      FC_W[1,12] := 0.07566059;
      FC_W[1,13] := 0.35968998;
      FC_W[1,14] := -0.17466193;
      FC_W[1,15] := 1.00617445;
      FC_W[1,16] := 0.29971626;
      FC_W[1,17] := -0.15427162;
      FC_W[1,18] := 0.06198071;
      FC_W[1,19] := 0.48209724;
      FC_W[1,20] := -1.77777910;
      FC_W[1,21] := 0.30678549;
      FC_W[1,22] := -0.06820694;
      FC_W[1,23] := -1.06389523;
      FC_W[1,24] := 1.40704405;
      FC_W[1,25] := 0.86564183;
      FC_W[1,26] := 0.86175865;
      FC_W[1,27] := -0.30832738;
      FC_W[1,28] := 0.12632002;
      FC_W[1,29] := 0.22659495;
      FC_W[1,30] := -0.13902418;
      FC_W[1,31] := -0.99291939;
      FC_W[2,0] := 0.04160358;
      FC_W[2,1] := 0.28197494;
      FC_W[2,2] := -0.02089060;
      FC_W[2,3] := 0.47015443;
      FC_W[2,4] := 0.34037617;
      FC_W[2,5] := -0.41242811;
      FC_W[2,6] := -0.82493418;
      FC_W[2,7] := 0.78098351;
      FC_W[2,8] := -0.39970401;
      FC_W[2,9] := 1.02419770;
      FC_W[2,10] := -0.33057141;
      FC_W[2,11] := 0.13100362;
      FC_W[2,12] := -1.50004947;
      FC_W[2,13] := -0.18024392;
      FC_W[2,14] := 0.19656396;
      FC_W[2,15] := -1.08431160;
      FC_W[2,16] := -0.22757976;
      FC_W[2,17] := -0.09310954;
      FC_W[2,18] := 1.20083344;
      FC_W[2,19] := -0.90194166;
      FC_W[2,20] := 0.46690372;
      FC_W[2,21] := -0.28373122;
      FC_W[2,22] := 0.44820097;
      FC_W[2,23] := 1.57939780;
      FC_W[2,24] := -0.41811836;
      FC_W[2,25] := 0.45971355;
      FC_W[2,26] := -0.05362111;
      FC_W[2,27] := -0.62090284;
      FC_W[2,28] := -0.41635084;
      FC_W[2,29] := 1.19535244;
      FC_W[2,30] := 0.22620986;
      FC_W[2,31] := -0.29096127;
      FC_W[3,0] := 0.69258898;
      FC_W[3,1] := -0.10189002;
      FC_W[3,2] := -0.35127911;
      FC_W[3,3] := -0.06208733;
      FC_W[3,4] := -0.31526309;
      FC_W[3,5] := -0.58414000;
      FC_W[3,6] := 0.04904716;
      FC_W[3,7] := 0.37988806;
      FC_W[3,8] := -0.33488220;
      FC_W[3,9] := 0.67849815;
      FC_W[3,10] := 0.02032584;
      FC_W[3,11] := -0.11450892;
      FC_W[3,12] := 0.75389469;
      FC_W[3,13] := -0.00020683;
      FC_W[3,14] := 0.11827329;
      FC_W[3,15] := 0.03889267;
      FC_W[3,16] := 0.17466927;
      FC_W[3,17] := -0.05837984;
      FC_W[3,18] := 0.16143340;
      FC_W[3,19] := -0.25548884;
      FC_W[3,20] := 0.36278751;
      FC_W[3,21] := 0.31648728;
      FC_W[3,22] := -0.78370738;
      FC_W[3,23] := -0.28512084;
      FC_W[3,24] := -0.33843708;
      FC_W[3,25] := 0.04330043;
      FC_W[3,26] := -0.25837252;
      FC_W[3,27] := 0.40221891;
      FC_W[3,28] := 0.07115368;
      FC_W[3,29] := 1.57388341;
      FC_W[3,30] := 0.08364432;
      FC_W[3,31] := 0.69666040;
      FC_W[4,0] := 0.17098659;
      FC_W[4,1] := 0.70854473;
      FC_W[4,2] := 0.32589009;
      FC_W[4,3] := -0.19657923;
      FC_W[4,4] := 0.02836942;
      FC_W[4,5] := -0.33067968;
      FC_W[4,6] := -0.28083199;
      FC_W[4,7] := 0.21882291;
      FC_W[4,8] := 0.44031367;
      FC_W[4,9] := -0.08098698;
      FC_W[4,10] := 0.40485817;
      FC_W[4,11] := -0.28698298;
      FC_W[4,12] := 0.25233796;
      FC_W[4,13] := -0.10523839;
      FC_W[4,14] := -0.44006598;
      FC_W[4,15] := -0.39039072;
      FC_W[4,16] := 0.15023036;
      FC_W[4,17] := 0.09987778;
      FC_W[4,18] := -0.55138695;
      FC_W[4,19] := 0.97002214;
      FC_W[4,20] := -1.32036424;
      FC_W[4,21] := 0.12111247;
      FC_W[4,22] := 0.17146327;
      FC_W[4,23] := -0.14426313;
      FC_W[4,24] := -1.44331551;
      FC_W[4,25] := -0.32387802;
      FC_W[4,26] := -0.86985487;
      FC_W[4,27] := 0.16190216;
      FC_W[4,28] := -0.25917780;
      FC_W[4,29] := 0.87935007;
      FC_W[4,30] := -0.04532806;
      FC_W[4,31] := 0.12371654;
      FC_W[5,0] := 0.16069181;
      FC_W[5,1] := 1.64132881;
      FC_W[5,2] := 0.09314496;
      FC_W[5,3] := 0.30746382;
      FC_W[5,4] := -0.44713461;
      FC_W[5,5] := -0.17269248;
      FC_W[5,6] := -0.43764487;
      FC_W[5,7] := -0.55917907;
      FC_W[5,8] := 0.07907125;
      FC_W[5,9] := 0.32444280;
      FC_W[5,10] := 0.17686915;
      FC_W[5,11] := -0.43060029;
      FC_W[5,12] := -0.11524609;
      FC_W[5,13] := -0.43634474;
      FC_W[5,14] := -0.84067672;
      FC_W[5,15] := 0.12469457;
      FC_W[5,16] := 0.36836424;
      FC_W[5,17] := -0.39146784;
      FC_W[5,18] := 0.77493954;
      FC_W[5,19] := -0.39445737;
      FC_W[5,20] := 0.13570420;
      FC_W[5,21] := -0.30796599;
      FC_W[5,22] := 0.57390678;
      FC_W[5,23] := -0.10128630;
      FC_W[5,24] := 0.46898919;
      FC_W[5,25] := -0.44309253;
      FC_W[5,26] := 0.08969644;
      FC_W[5,27] := -0.19782862;
      FC_W[5,28] := 2.73940182;
      FC_W[5,29] := 0.16153421;
      FC_W[5,30] := -0.12013239;
      FC_W[5,31] := -0.56593496;
      FC_W[6,0] := -0.57114196;
      FC_W[6,1] := 1.38476813;
      FC_W[6,2] := 1.11997521;
      FC_W[6,3] := 0.02632367;
      FC_W[6,4] := -0.45034066;
      FC_W[6,5] := 1.03288424;
      FC_W[6,6] := -0.40567783;
      FC_W[6,7] := 0.16608752;
      FC_W[6,8] := 0.03270433;
      FC_W[6,9] := -0.35795641;
      FC_W[6,10] := 0.00975101;
      FC_W[6,11] := -0.41937128;
      FC_W[6,12] := -0.19609804;
      FC_W[6,13] := -0.28889647;
      FC_W[6,14] := -0.96404856;
      FC_W[6,15] := 0.08155423;
      FC_W[6,16] := 0.09745946;
      FC_W[6,17] := 0.17013049;
      FC_W[6,18] := 0.17057557;
      FC_W[6,19] := -0.79009062;
      FC_W[6,20] := 0.26148456;
      FC_W[6,21] := -0.41126329;
      FC_W[6,22] := -0.92280918;
      FC_W[6,23] := -0.19497190;
      FC_W[6,24] := 0.56321335;
      FC_W[6,25] := -0.69397563;
      FC_W[6,26] := -0.11093070;
      FC_W[6,27] := -0.12486640;
      FC_W[6,28] := -0.51809597;
      FC_W[6,29] := 0.44581598;
      FC_W[6,30] := -0.07224379;
      FC_W[6,31] := 0.58158380;
      FC_W[7,0] := 0.41476303;
      FC_W[7,1] := -0.03894622;
      FC_W[7,2] := -0.50756085;
      FC_W[7,3] := -0.26348099;
      FC_W[7,4] := 0.08712668;
      FC_W[7,5] := -0.37651458;
      FC_W[7,6] := 0.26482788;
      FC_W[7,7] := -0.29581240;
      FC_W[7,8] := 0.05395310;
      FC_W[7,9] := 0.41241437;
      FC_W[7,10] := -0.15156971;
      FC_W[7,11] := 0.26749688;
      FC_W[7,12] := 0.97054368;
      FC_W[7,13] := -0.03540496;
      FC_W[7,14] := -0.09778718;
      FC_W[7,15] := -0.39193475;
      FC_W[7,16] := -0.01532598;
      FC_W[7,17] := -0.11887385;
      FC_W[7,18] := -0.30799413;
      FC_W[7,19] := -0.20951317;
      FC_W[7,20] := 0.46884289;
      FC_W[7,21] := 0.08239307;
      FC_W[7,22] := -0.41243985;
      FC_W[7,23] := -0.14386208;
      FC_W[7,24] := -0.56366146;
      FC_W[7,25] := 0.05347069;
      FC_W[7,26] := -0.06422243;
      FC_W[7,27] := -0.14232105;
      FC_W[7,28] := 0.08967300;
      FC_W[7,29] := 2.09215212;
      FC_W[7,30] := -0.41609016;
      FC_W[7,31] := 0.61930108;
      FC_W[8,0] := 0.41138357;
      FC_W[8,1] := -0.13876545;
      FC_W[8,2] := -0.47696707;
      FC_W[8,3] := -0.58067173;
      FC_W[8,4] := -0.76539934;
      FC_W[8,5] := -0.48228866;
      FC_W[8,6] := 0.25288635;
      FC_W[8,7] := 1.26393640;
      FC_W[8,8] := -0.18708183;
      FC_W[8,9] := 1.05916786;
      FC_W[8,10] := -0.21405555;
      FC_W[8,11] := -0.73763049;
      FC_W[8,12] := -0.49388906;
      FC_W[8,13] := 0.23774624;
      FC_W[8,14] := 0.03641314;
      FC_W[8,15] := 0.43136188;
      FC_W[8,16] := -0.34853166;
      FC_W[8,17] := 0.45351282;
      FC_W[8,18] := 0.12007232;
      FC_W[8,19] := -0.09311971;
      FC_W[8,20] := 0.10139518;
      FC_W[8,21] := 0.13798890;
      FC_W[8,22] := -0.75192511;
      FC_W[8,23] := -0.33668301;
      FC_W[8,24] := 0.14659424;
      FC_W[8,25] := -0.00453089;
      FC_W[8,26] := -0.35082975;
      FC_W[8,27] := 0.47500724;
      FC_W[8,28] := 0.02143906;
      FC_W[8,29] := 0.81066149;
      FC_W[8,30] := 0.42516547;
      FC_W[8,31] := 1.48935926;
      FC_W[9,0] := 0.29422590;
      FC_W[9,1] := -0.02413537;
      FC_W[9,2] := -0.57707560;
      FC_W[9,3] := -0.44330636;
      FC_W[9,4] := -0.02986326;
      FC_W[9,5] := -0.32138100;
      FC_W[9,6] := 0.33747303;
      FC_W[9,7] := -0.02603977;
      FC_W[9,8] := 0.16214876;
      FC_W[9,9] := 0.54148763;
      FC_W[9,10] := -0.23998420;
      FC_W[9,11] := 0.06466576;
      FC_W[9,12] := 0.47260144;
      FC_W[9,13] := 0.04922871;
      FC_W[9,14] := -0.13990949;
      FC_W[9,15] := -0.24958028;
      FC_W[9,16] := -0.20513535;
      FC_W[9,17] := 0.11604570;
      FC_W[9,18] := -0.38338530;
      FC_W[9,19] := -0.16188677;
      FC_W[9,20] := 0.37325716;
      FC_W[9,21] := -0.01747377;
      FC_W[9,22] := -0.37153879;
      FC_W[9,23] := -0.15362059;
      FC_W[9,24] := -0.37243831;
      FC_W[9,25] := 0.01588886;
      FC_W[9,26] := -0.08001896;
      FC_W[9,27] := -0.14023392;
      FC_W[9,28] := 0.07176708;
      FC_W[9,29] := 1.81881726;
      FC_W[9,30] := -0.30937484;
      FC_W[9,31] := 0.93038040;
      FC_W[10,0] := -0.05140001;
      FC_W[10,1] := -0.21192010;
      FC_W[10,2] := -0.34014732;
      FC_W[10,3] := -0.41698745;
      FC_W[10,4] := 1.15412712;
      FC_W[10,5] := -0.76638728;
      FC_W[10,6] := -0.36194009;
      FC_W[10,7] := -0.14446546;
      FC_W[10,8] := 0.05265777;
      FC_W[10,9] := 0.60072738;
      FC_W[10,10] := 0.43118945;
      FC_W[10,11] := 0.83294547;
      FC_W[10,12] := 0.67825025;
      FC_W[10,13] := 0.19051756;
      FC_W[10,14] := 1.69663048;
      FC_W[10,15] := -0.22305325;
      FC_W[10,16] := -0.32500228;
      FC_W[10,17] := 0.31870443;
      FC_W[10,18] := 0.10095058;
      FC_W[10,19] := -0.75147802;
      FC_W[10,20] := -0.45519939;
      FC_W[10,21] := 0.01013143;
      FC_W[10,22] := 0.00206094;
      FC_W[10,23] := 0.25191501;
      FC_W[10,24] := 0.39815706;
      FC_W[10,25] := -0.34215525;
      FC_W[10,26] := -0.22784939;
      FC_W[10,27] := 0.34508327;
      FC_W[10,28] := 1.05789781;
      FC_W[10,29] := 1.05650342;
      FC_W[10,30] := -0.25448412;
      FC_W[10,31] := 1.19635260;
      FC_W[11,0] := -0.60992318;
      FC_W[11,1] := 0.06451012;
      FC_W[11,2] := -0.06141585;
      FC_W[11,3] := 0.26182047;
      FC_W[11,4] := -0.30671248;
      FC_W[11,5] := -0.15614234;
      FC_W[11,6] := 0.20122612;
      FC_W[11,7] := -0.25060847;
      FC_W[11,8] := 0.21109147;
      FC_W[11,9] := 0.34703916;
      FC_W[11,10] := -1.65234506;
      FC_W[11,11] := -0.15922636;
      FC_W[11,12] := -0.04707455;
      FC_W[11,13] := 0.20130210;
      FC_W[11,14] := -0.29188156;
      FC_W[11,15] := 1.00682425;
      FC_W[11,16] := 1.30854654;
      FC_W[11,17] := 0.41931316;
      FC_W[11,18] := 0.32618555;
      FC_W[11,19] := -0.02777285;
      FC_W[11,20] := -0.33175266;
      FC_W[11,21] := -0.60335326;
      FC_W[11,22] := 0.34577838;
      FC_W[11,23] := 0.24502832;
      FC_W[11,24] := 0.50228852;
      FC_W[11,25] := -0.19970542;
      FC_W[11,26] := 0.01159031;
      FC_W[11,27] := 0.17553034;
      FC_W[11,28] := -0.36863360;
      FC_W[11,29] := 0.21139398;
      FC_W[11,30] := 0.41804573;
      FC_W[11,31] := 0.16023155;
      FC_W[12,0] := 0.16499591;
      FC_W[12,1] := 0.14349781;
      FC_W[12,2] := -0.01990420;
      FC_W[12,3] := 0.96575189;
      FC_W[12,4] := -0.45016506;
      FC_W[12,5] := -0.58705819;
      FC_W[12,6] := -0.48950329;
      FC_W[12,7] := -0.19916040;
      FC_W[12,8] := 0.57504302;
      FC_W[12,9] := 0.15542965;
      FC_W[12,10] := -0.41850585;
      FC_W[12,11] := -0.14737980;
      FC_W[12,12] := 0.29411027;
      FC_W[12,13] := 0.31234270;
      FC_W[12,14] := -0.10017619;
      FC_W[12,15] := 1.20768833;
      FC_W[12,16] := 1.27741170;
      FC_W[12,17] := -0.28955090;
      FC_W[12,18] := 0.87563890;
      FC_W[12,19] := -0.36919677;
      FC_W[12,20] := -0.45485532;
      FC_W[12,21] := -0.81351525;
      FC_W[12,22] := 0.01215564;
      FC_W[12,23] := 0.66354555;
      FC_W[12,24] := 0.64124012;
      FC_W[12,25] := -0.36083624;
      FC_W[12,26] := -0.03435243;
      FC_W[12,27] := 0.60670197;
      FC_W[12,28] := -0.31781450;
      FC_W[12,29] := 0.27313688;
      FC_W[12,30] := 0.53784895;
      FC_W[12,31] := -0.24992017;
      FC_W[13,0] := 1.15009689;
      FC_W[13,1] := 0.24936195;
      FC_W[13,2] := -0.18515313;
      FC_W[13,3] := 0.81901830;
      FC_W[13,4] := -0.05867874;
      FC_W[13,5] := -0.56633902;
      FC_W[13,6] := 0.23188661;
      FC_W[13,7] := 0.06102761;
      FC_W[13,8] := -0.12947020;
      FC_W[13,9] := -0.30986655;
      FC_W[13,10] := -0.05449111;
      FC_W[13,11] := 0.41703042;
      FC_W[13,12] := -0.64008683;
      FC_W[13,13] := -0.47276545;
      FC_W[13,14] := 0.17531119;
      FC_W[13,15] := -1.03741860;
      FC_W[13,16] := 0.60905075;
      FC_W[13,17] := -0.09274173;
      FC_W[13,18] := -0.27676162;
      FC_W[13,19] := 0.67100716;
      FC_W[13,20] := -0.97478300;
      FC_W[13,21] := 0.11877309;
      FC_W[13,22] := 0.60747856;
      FC_W[13,23] := -0.10786309;
      FC_W[13,24] := -0.19802028;
      FC_W[13,25] := -1.18054771;
      FC_W[13,26] := 2.67729783;
      FC_W[13,27] := 0.40492588;
      FC_W[13,28] := -0.12357215;
      FC_W[13,29] := 0.05446408;
      FC_W[13,30] := -0.33658338;
      FC_W[13,31] := -0.28736502;
      FC_W[14,0] := -1.09515917;
      FC_W[14,1] := -0.22429042;
      FC_W[14,2] := -1.36213231;
      FC_W[14,3] := 1.22893906;
      FC_W[14,4] := 0.23815246;
      FC_W[14,5] := -1.80320215;
      FC_W[14,6] := 0.25902322;
      FC_W[14,7] := 1.75334704;
      FC_W[14,8] := 2.21751308;
      FC_W[14,9] := -1.82321739;
      FC_W[14,10] := -1.16461563;
      FC_W[14,11] := -0.11827917;
      FC_W[14,12] := 0.38857111;
      FC_W[14,13] := 0.05780562;
      FC_W[14,14] := -1.02024376;
      FC_W[14,15] := 0.64406765;
      FC_W[14,16] := -1.86519647;
      FC_W[14,17] := 0.51558846;
      FC_W[14,18] := 0.29011348;
      FC_W[14,19] := -1.91969121;
      FC_W[14,20] := 0.18231264;
      FC_W[14,21] := 2.35030413;
      FC_W[14,22] := 0.28205252;
      FC_W[14,23] := -0.05250929;
      FC_W[14,24] := 0.08201724;
      FC_W[14,25] := -2.43822980;
      FC_W[14,26] := -0.05353496;
      FC_W[14,27] := -0.08439671;
      FC_W[14,28] := 0.31032041;
      FC_W[14,29] := -0.01394748;
      FC_W[14,30] := 0.17681596;
      FC_W[14,31] := -1.01465368;
      FC_W[15,0] := -0.76047558;
      FC_W[15,1] := 0.18870419;
      FC_W[15,2] := -0.05700897;
      FC_W[15,3] := -0.52280545;
      FC_W[15,4] := 0.75352377;
      FC_W[15,5] := 0.28025728;
      FC_W[15,6] := -0.01245948;
      FC_W[15,7] := 0.32771844;
      FC_W[15,8] := -0.20845552;
      FC_W[15,9] := -0.46889994;
      FC_W[15,10] := -1.00782621;
      FC_W[15,11] := -0.25399303;
      FC_W[15,12] := 0.32204163;
      FC_W[15,13] := -0.28043103;
      FC_W[15,14] := -0.12425613;
      FC_W[15,15] := 0.16964360;
      FC_W[15,16] := 1.18621874;
      FC_W[15,17] := 0.55311561;
      FC_W[15,18] := 1.06978226;
      FC_W[15,19] := 0.18990995;
      FC_W[15,20] := 0.48186046;
      FC_W[15,21] := -0.44492897;
      FC_W[15,22] := 0.25515074;
      FC_W[15,23] := -1.14194119;
      FC_W[15,24] := -0.87563568;
      FC_W[15,25] := 0.54568601;
      FC_W[15,26] := 0.49307632;
      FC_W[15,27] := 0.92335260;
      FC_W[15,28] := -0.08592582;
      FC_W[15,29] := 0.41658750;
      FC_W[15,30] := 2.08434486;
      FC_W[15,31] := -0.23699243;
      FC_W[16,0] := 0.45081332;
      FC_W[16,1] := 0.21935241;
      FC_W[16,2] := 0.10121434;
      FC_W[16,3] := -0.55789620;
      FC_W[16,4] := 0.45296088;
      FC_W[16,5] := 0.34732810;
      FC_W[16,6] := 1.75819397;
      FC_W[16,7] := -0.05926482;
      FC_W[16,8] := 0.96878350;
      FC_W[16,9] := 0.08046997;
      FC_W[16,10] := 0.37100121;
      FC_W[16,11] := -0.28692111;
      FC_W[16,12] := 0.01441160;
      FC_W[16,13] := -0.00036847;
      FC_W[16,14] := 0.08188357;
      FC_W[16,15] := -0.76726955;
      FC_W[16,16] := 0.58374065;
      FC_W[16,17] := -0.63479686;
      FC_W[16,18] := -2.68864226;
      FC_W[16,19] := -0.27776572;
      FC_W[16,20] := -0.24950075;
      FC_W[16,21] := 1.06383419;
      FC_W[16,22] := -1.58518887;
      FC_W[16,23] := 3.18674827;
      FC_W[16,24] := 0.32398152;
      FC_W[16,25] := 0.74144083;
      FC_W[16,26] := -0.01374951;
      FC_W[16,27] := 1.09727502;
      FC_W[16,28] := 0.24661481;
      FC_W[16,29] := -0.21010247;
      FC_W[16,30] := 1.18042016;
      FC_W[16,31] := -0.61184710;
      FC_W[17,0] := -0.16353357;
      FC_W[17,1] := -0.69889224;
      FC_W[17,2] := -0.67269742;
      FC_W[17,3] := -1.10959411;
      FC_W[17,4] := 0.66946703;
      FC_W[17,5] := -0.88466114;
      FC_W[17,6] := 1.81482458;
      FC_W[17,7] := 0.85526884;
      FC_W[17,8] := -0.42613694;
      FC_W[17,9] := -1.93829262;
      FC_W[17,10] := 2.12208724;
      FC_W[17,11] := 0.87851965;
      FC_W[17,12] := -1.60542023;
      FC_W[17,13] := -0.39448434;
      FC_W[17,14] := -0.57687348;
      FC_W[17,15] := -0.18362631;
      FC_W[17,16] := 2.05336404;
      FC_W[17,17] := -0.54798490;
      FC_W[17,18] := 0.09048657;
      FC_W[17,19] := -1.08607030;
      FC_W[17,20] := 0.51026022;
      FC_W[17,21] := -0.92757076;
      FC_W[17,22] := -0.97661769;
      FC_W[17,23] := -0.05264290;
      FC_W[17,24] := -0.09709509;
      FC_W[17,25] := -1.65425158;
      FC_W[17,26] := -0.74785799;
      FC_W[17,27] := 0.17301857;
      FC_W[17,28] := 0.38459933;
      FC_W[17,29] := 0.64529657;
      FC_W[17,30] := -2.37725043;
      FC_W[17,31] := -0.66769147;
      FC_W[18,0] := -0.58205122;
      FC_W[18,1] := 0.17416364;
      FC_W[18,2] := -0.21704014;
      FC_W[18,3] := -0.15796715;
      FC_W[18,4] := -0.06134655;
      FC_W[18,5] := 0.18992065;
      FC_W[18,6] := -0.55935055;
      FC_W[18,7] := -1.69722903;
      FC_W[18,8] := -0.16580440;
      FC_W[18,9] := -0.49130309;
      FC_W[18,10] := -0.70880896;
      FC_W[18,11] := 0.16293578;
      FC_W[18,12] := -2.99989247;
      FC_W[18,13] := -0.07632764;
      FC_W[18,14] := -0.36394569;
      FC_W[18,15] := 2.71546102;
      FC_W[18,16] := -1.11394608;
      FC_W[18,17] := 0.23080237;
      FC_W[18,18] := 0.42428958;
      FC_W[18,19] := -0.31673199;
      FC_W[18,20] := 0.35938102;
      FC_W[18,21] := -0.28474978;
      FC_W[18,22] := 0.23496971;
      FC_W[18,23] := -0.56855541;
      FC_W[18,24] := 0.13188744;
      FC_W[18,25] := 0.08833195;
      FC_W[18,26] := -0.28358048;
      FC_W[18,27] := 2.70895100;
      FC_W[18,28] := -0.37571719;
      FC_W[18,29] := 2.44771218;
      FC_W[18,30] := 1.01540816;
      FC_W[18,31] := -0.99419475;
      FC_W[19,0] := -0.04479429;
      FC_W[19,1] := -0.03746313;
      FC_W[19,2] := -0.13186198;
      FC_W[19,3] := 0.34855995;
      FC_W[19,4] := 0.02845483;
      FC_W[19,5] := -0.42788455;
      FC_W[19,6] := 0.28289452;
      FC_W[19,7] := 0.42844373;
      FC_W[19,8] := 0.57057315;
      FC_W[19,9] := -0.34337267;
      FC_W[19,10] := -0.41033122;
      FC_W[19,11] := -0.18694647;
      FC_W[19,12] := 0.05562596;
      FC_W[19,13] := 0.04664620;
      FC_W[19,14] := -0.08783104;
      FC_W[19,15] := 0.16602120;
      FC_W[19,16] := -0.26911020;
      FC_W[19,17] := 0.21557054;
      FC_W[19,18] := 0.10632721;
      FC_W[19,19] := -0.38928598;
      FC_W[19,20] := -0.12570058;
      FC_W[19,21] := -2.12742734;
      FC_W[19,22] := -0.22360966;
      FC_W[19,23] := -0.23273115;
      FC_W[19,24] := 0.03732495;
      FC_W[19,25] := -0.41173750;
      FC_W[19,26] := 0.04321238;
      FC_W[19,27] := -0.09780092;
      FC_W[19,28] := 0.07972930;
      FC_W[19,29] := -0.04350290;
      FC_W[19,30] := 0.34195364;
      FC_W[19,31] := -0.30817261;
      FC_W[20,0] := 0.83343393;
      FC_W[20,1] := 0.58159441;
      FC_W[20,2] := -0.54344225;
      FC_W[20,3] := 0.15104640;
      FC_W[20,4] := 0.51991045;
      FC_W[20,5] := -0.79415458;
      FC_W[20,6] := 1.20831060;
      FC_W[20,7] := 0.07056488;
      FC_W[20,8] := 0.07098699;
      FC_W[20,9] := 0.00417417;
      FC_W[20,10] := 0.01662889;
      FC_W[20,11] := 0.43986788;
      FC_W[20,12] := 0.04565306;
      FC_W[20,13] := 0.36652237;
      FC_W[20,14] := 1.53537381;
      FC_W[20,15] := 0.13102606;
      FC_W[20,16] := -0.04194741;
      FC_W[20,17] := 0.24626848;
      FC_W[20,18] := -0.06461809;
      FC_W[20,19] := 0.41678023;
      FC_W[20,20] := 0.11291907;
      FC_W[20,21] := 0.58736563;
      FC_W[20,22] := 0.37338239;
      FC_W[20,23] := -0.43781069;
      FC_W[20,24] := -0.26015314;
      FC_W[20,25] := 0.77599698;
      FC_W[20,26] := -0.25086293;
      FC_W[20,27] := 0.14930426;
      FC_W[20,28] := -0.29598835;
      FC_W[20,29] := -0.65816528;
      FC_W[20,30] := -0.29212403;
      FC_W[20,31] := -0.35731244;
      FC_W[21,0] := -0.78355730;
      FC_W[21,1] := -0.09190790;
      FC_W[21,2] := 2.04684353;
      FC_W[21,3] := -0.52632159;
      FC_W[21,4] := 0.00004623;
      FC_W[21,5] := -0.41394150;
      FC_W[21,6] := 0.00152126;
      FC_W[21,7] := -0.09166983;
      FC_W[21,8] := 0.22487646;
      FC_W[21,9] := 0.55625015;
      FC_W[21,10] := 0.45326176;
      FC_W[21,11] := -0.36226249;
      FC_W[21,12] := 0.35516575;
      FC_W[21,13] := 1.12550521;
      FC_W[21,14] := -0.56490552;
      FC_W[21,15] := 0.29733366;
      FC_W[21,16] := -0.13095240;
      FC_W[21,17] := -0.62664920;
      FC_W[21,18] := -0.68398547;
      FC_W[21,19] := -0.36049438;
      FC_W[21,20] := 0.76424283;
      FC_W[21,21] := 0.14176156;
      FC_W[21,22] := 0.17250934;
      FC_W[21,23] := -0.62825954;
      FC_W[21,24] := -0.29867983;
      FC_W[21,25] := -0.32782140;
      FC_W[21,26] := -0.11939523;
      FC_W[21,27] := -0.13114350;
      FC_W[21,28] := -0.02881289;
      FC_W[21,29] := 0.40359056;
      FC_W[21,30] := 0.24945424;
      FC_W[21,31] := 0.11648370;
      FC_W[22,0] := 1.11175954;
      FC_W[22,1] := 0.34547076;
      FC_W[22,2] := 0.14727411;
      FC_W[22,3] := 0.63355762;
      FC_W[22,4] := 1.23095477;
      FC_W[22,5] := 0.22958253;
      FC_W[22,6] := -0.27086827;
      FC_W[22,7] := 0.21812293;
      FC_W[22,8] := 0.34522176;
      FC_W[22,9] := -0.30138829;
      FC_W[22,10] := -0.11115979;
      FC_W[22,11] := -0.99961066;
      FC_W[22,12] := -0.28910354;
      FC_W[22,13] := -0.28956577;
      FC_W[22,14] := -0.04969905;
      FC_W[22,15] := -0.22805935;
      FC_W[22,16] := 0.68084496;
      FC_W[22,17] := -0.59066468;
      FC_W[22,18] := -0.91510123;
      FC_W[22,19] := 0.36468261;
      FC_W[22,20] := 0.44435018;
      FC_W[22,21] := -0.09364665;
      FC_W[22,22] := 0.29944962;
      FC_W[22,23] := -0.92394197;
      FC_W[22,24] := 0.02677452;
      FC_W[22,25] := -1.25928640;
      FC_W[22,26] := -0.08920673;
      FC_W[22,27] := -0.22473238;
      FC_W[22,28] := -0.18966107;
      FC_W[22,29] := -0.15222032;
      FC_W[22,30] := 0.28112322;
      FC_W[22,31] := 0.07603560;
      FC_W[23,0] := 0.94918245;
      FC_W[23,1] := -0.16944362;
      FC_W[23,2] := -0.64516091;
      FC_W[23,3] := 0.01417535;
      FC_W[23,4] := 1.17094791;
      FC_W[23,5] := -0.46294600;
      FC_W[23,6] := 0.63886625;
      FC_W[23,7] := 0.59459019;
      FC_W[23,8] := -1.25560164;
      FC_W[23,9] := -0.41550717;
      FC_W[23,10] := -0.89923918;
      FC_W[23,11] := -2.04026842;
      FC_W[23,12] := 0.38108230;
      FC_W[23,13] := -0.46252671;
      FC_W[23,14] := 0.36853698;
      FC_W[23,15] := -0.68918151;
      FC_W[23,16] := 0.25558072;
      FC_W[23,17] := -0.33933294;
      FC_W[23,18] := -0.42984211;
      FC_W[23,19] := -0.58996665;
      FC_W[23,20] := -0.85563028;
      FC_W[23,21] := -0.00377321;
      FC_W[23,22] := 0.30137330;
      FC_W[23,23] := 0.55249846;
      FC_W[23,24] := 0.67464733;
      FC_W[23,25] := 0.68203866;
      FC_W[23,26] := 1.75322306;
      FC_W[23,27] := 0.65638542;
      FC_W[23,28] := -0.60190219;
      FC_W[23,29] := -0.19525060;
      FC_W[23,30] := -1.64320982;
      FC_W[23,31] := 0.09680892;
      FC_W[24,0] := 1.70816791;
      FC_W[24,1] := 0.19184691;
      FC_W[24,2] := 0.43070525;
      FC_W[24,3] := 0.47347856;
      FC_W[24,4] := 1.06446636;
      FC_W[24,5] := 0.82846808;
      FC_W[24,6] := -0.14924394;
      FC_W[24,7] := 0.48391837;
      FC_W[24,8] := 0.10338319;
      FC_W[24,9] := -0.42541158;
      FC_W[24,10] := -0.46907026;
      FC_W[24,11] := -1.26659918;
      FC_W[24,12] := 0.00209635;
      FC_W[24,13] := -0.58223796;
      FC_W[24,14] := 0.35529405;
      FC_W[24,15] := -0.17281178;
      FC_W[24,16] := 0.78266329;
      FC_W[24,17] := -0.47265151;
      FC_W[24,18] := -0.52031809;
      FC_W[24,19] := 0.60595226;
      FC_W[24,20] := 0.93959928;
      FC_W[24,21] := -0.07003678;
      FC_W[24,22] := 0.40464661;
      FC_W[24,23] := -0.47159809;
      FC_W[24,24] := -0.21403076;
      FC_W[24,25] := -1.99785328;
      FC_W[24,26] := -0.31490597;
      FC_W[24,27] := 0.22405344;
      FC_W[24,28] := -0.12689462;
      FC_W[24,29] := -0.13865131;
      FC_W[24,30] := 0.19015649;
      FC_W[24,31] := -0.10777009;
      FC_W[25,0] := 1.68829179;
      FC_W[25,1] := 0.20417857;
      FC_W[25,2] := 0.41045186;
      FC_W[25,3] := 0.49043059;
      FC_W[25,4] := 1.10725451;
      FC_W[25,5] := 0.79095447;
      FC_W[25,6] := -0.15897395;
      FC_W[25,7] := 0.44460773;
      FC_W[25,8] := 0.12746778;
      FC_W[25,9] := -0.38992313;
      FC_W[25,10] := -0.42752251;
      FC_W[25,11] := -1.26661718;
      FC_W[25,12] := -0.01255040;
      FC_W[25,13] := -0.56674266;
      FC_W[25,14] := 0.30763030;
      FC_W[25,15] := -0.16670777;
      FC_W[25,16] := 0.78490394;
      FC_W[25,17] := -0.41297758;
      FC_W[25,18] := -0.56244904;
      FC_W[25,19] := 0.59661794;
      FC_W[25,20] := 0.91377634;
      FC_W[25,21] := -0.07476726;
      FC_W[25,22] := 0.39158839;
      FC_W[25,23] := -0.50374097;
      FC_W[25,24] := -0.20792229;
      FC_W[25,25] := -1.98061037;
      FC_W[25,26] := -0.29893139;
      FC_W[25,27] := 0.20798860;
      FC_W[25,28] := -0.13327917;
      FC_W[25,29] := -0.14427565;
      FC_W[25,30] := 0.18739435;
      FC_W[25,31] := -0.12663475;
      FC_W[26,0] := 2.09756184;
      FC_W[26,1] := 0.30979156;
      FC_W[26,2] := -0.93082160;
      FC_W[26,3] := 1.12418640;
      FC_W[26,4] := -0.21458086;
      FC_W[26,5] := -0.20711824;
      FC_W[26,6] := 0.13515653;
      FC_W[26,7] := -0.10551527;
      FC_W[26,8] := -0.78610575;
      FC_W[26,9] := -0.74051434;
      FC_W[26,10] := -0.11710767;
      FC_W[26,11] := 0.56832963;
      FC_W[26,12] := -0.63929403;
      FC_W[26,13] := -0.61865294;
      FC_W[26,14] := -0.03843753;
      FC_W[26,15] := -0.58638787;
      FC_W[26,16] := 0.65063626;
      FC_W[26,17] := 0.77623236;
      FC_W[26,18] := -1.90139818;
      FC_W[26,19] := -0.35095820;
      FC_W[26,20] := -0.92717338;
      FC_W[26,21] := -0.01369499;
      FC_W[26,22] := 0.80340147;
      FC_W[26,23] := -0.95347393;
      FC_W[26,24] := 0.83274955;
      FC_W[26,25] := -0.80403948;
      FC_W[26,26] := 0.11611202;
      FC_W[26,27] := -0.82351989;
      FC_W[26,28] := -0.07890483;
      FC_W[26,29] := -0.10332011;
      FC_W[26,30] := 0.82299954;
      FC_W[26,31] := -0.11604206;
      FC_W[27,0] := -0.21567799;
      FC_W[27,1] := -0.17982188;
      FC_W[27,2] := 1.61042237;
      FC_W[27,3] := -0.04066473;
      FC_W[27,4] := 0.35580903;
      FC_W[27,5] := 0.17180133;
      FC_W[27,6] := -0.03739715;
      FC_W[27,7] := 0.47538793;
      FC_W[27,8] := 0.08444246;
      FC_W[27,9] := -0.20834255;
      FC_W[27,10] := -0.25132874;
      FC_W[27,11] := -0.09292793;
      FC_W[27,12] := 0.09512535;
      FC_W[27,13] := 1.73640633;
      FC_W[27,14] := -0.84270179;
      FC_W[27,15] := 0.10921801;
      FC_W[27,16] := 0.14793324;
      FC_W[27,17] := 0.00623075;
      FC_W[27,18] := -0.40309554;
      FC_W[27,19] := -0.10969527;
      FC_W[27,20] := 0.62004441;
      FC_W[27,21] := -0.05732905;
      FC_W[27,22] := 0.31839165;
      FC_W[27,23] := 0.20006965;
      FC_W[27,24] := -0.76557893;
      FC_W[27,25] := 0.08809149;
      FC_W[27,26] := -0.23099069;
      FC_W[27,27] := 0.52423984;
      FC_W[27,28] := 0.15881240;
      FC_W[27,29] := 0.15915051;
      FC_W[27,30] := -0.01910155;
      FC_W[27,31] := 0.50223130;
      FC_W[28,0] := 0.38221422;
      FC_W[28,1] := 0.00505643;
      FC_W[28,2] := 0.47086298;
      FC_W[28,3] := 0.38442624;
      FC_W[28,4] := -0.36451018;
      FC_W[28,5] := 0.23073554;
      FC_W[28,6] := 0.58682746;
      FC_W[28,7] := -0.31383422;
      FC_W[28,8] := 0.26966298;
      FC_W[28,9] := 0.52483726;
      FC_W[28,10] := -0.34839612;
      FC_W[28,11] := -0.04066939;
      FC_W[28,12] := 0.00757548;
      FC_W[28,13] := -0.89035267;
      FC_W[28,14] := -0.37031823;
      FC_W[28,15] := -0.28977558;
      FC_W[28,16] := 0.20845301;
      FC_W[28,17] := -0.68783289;
      FC_W[28,18] := 0.18428198;
      FC_W[28,19] := -1.10686350;
      FC_W[28,20] := -0.96242166;
      FC_W[28,21] := 0.16471045;
      FC_W[28,22] := -0.18428743;
      FC_W[28,23] := -0.42145190;
      FC_W[28,24] := -1.93459392;
      FC_W[28,25] := -0.20813486;
      FC_W[28,26] := -0.20319073;
      FC_W[28,27] := 0.50201613;
      FC_W[28,28] := -0.07826387;
      FC_W[28,29] := -0.16438225;
      FC_W[28,30] := -0.21372633;
      FC_W[28,31] := 0.31741613;
      FC_W[29,0] := 0.64168429;
      FC_W[29,1] := 0.44630602;
      FC_W[29,2] := -0.78172582;
      FC_W[29,3] := -0.80917108;
      FC_W[29,4] := 2.00600052;
      FC_W[29,5] := -0.28020853;
      FC_W[29,6] := 0.47931615;
      FC_W[29,7] := -1.29415607;
      FC_W[29,8] := 0.46214828;
      FC_W[29,9] := 2.15377712;
      FC_W[29,10] := 2.74666047;
      FC_W[29,11] := -0.29106671;
      FC_W[29,12] := 0.74129343;
      FC_W[29,13] := -0.13792343;
      FC_W[29,14] := -2.72200084;
      FC_W[29,15] := 0.92555773;
      FC_W[29,16] := -1.05131578;
      FC_W[29,17] := 3.75333142;
      FC_W[29,18] := 0.45929980;
      FC_W[29,19] := 0.72067416;
      FC_W[29,20] := 0.08021349;
      FC_W[29,21] := 0.19734156;
      FC_W[29,22] := 0.97599524;
      FC_W[29,23] := 0.68264025;
      FC_W[29,24] := 0.16812357;
      FC_W[29,25] := -1.16828287;
      FC_W[29,26] := 0.26183292;
      FC_W[29,27] := 1.09284210;
      FC_W[29,28] := -0.32955399;
      FC_W[29,29] := -0.92582864;
      FC_W[29,30] := -0.27071735;
      FC_W[29,31] := -1.27781820;
      FC_W[30,0] := 1.10601306;
      FC_W[30,1] := 0.35029322;
      FC_W[30,2] := 0.14326763;
      FC_W[30,3] := 0.63553667;
      FC_W[30,4] := 1.23359120;
      FC_W[30,5] := 0.22257970;
      FC_W[30,6] := -0.26709387;
      FC_W[30,7] := 0.21314621;
      FC_W[30,8] := 0.34742895;
      FC_W[30,9] := -0.29764310;
      FC_W[30,10] := -0.10436807;
      FC_W[30,11] := -0.99244106;
      FC_W[30,12] := -0.29116562;
      FC_W[30,13] := -0.28640470;
      FC_W[30,14] := -0.05612181;
      FC_W[30,15] := -0.22917078;
      FC_W[30,16] := 0.67629182;
      FC_W[30,17] := -0.59625685;
      FC_W[30,18] := -0.91921037;
      FC_W[30,19] := 0.36291701;
      FC_W[30,20] := 0.43871662;
      FC_W[30,21] := -0.09457398;
      FC_W[30,22] := 0.30445847;
      FC_W[30,23] := -0.92936188;
      FC_W[30,24] := 0.02971039;
      FC_W[30,25] := -1.25080836;
      FC_W[30,26] := -0.08806182;
      FC_W[30,27] := -0.23112479;
      FC_W[30,28] := -0.19110020;
      FC_W[30,29] := -0.15325592;
      FC_W[30,30] := 0.28191712;
      FC_W[30,31] := 0.07912993;
      FC_W[31,0] := 1.12223732;
      FC_W[31,1] := 0.36431006;
      FC_W[31,2] := 0.46958429;
      FC_W[31,3] := 1.85451174;
      FC_W[31,4] := 1.60030389;
      FC_W[31,5] := -0.15342215;
      FC_W[31,6] := 0.42601490;
      FC_W[31,7] := 0.20544830;
      FC_W[31,8] := -0.83132565;
      FC_W[31,9] := -0.26838920;
      FC_W[31,10] := -0.80358034;
      FC_W[31,11] := -0.01014836;
      FC_W[31,12] := -0.12229779;
      FC_W[31,13] := -0.43185377;
      FC_W[31,14] := -0.42969078;
      FC_W[31,15] := -0.43150717;
      FC_W[31,16] := 0.37160653;
      FC_W[31,17] := -1.10086751;
      FC_W[31,18] := -0.93033099;
      FC_W[31,19] := 0.68914485;
      FC_W[31,20] := 0.25832367;
      FC_W[31,21] := -0.17015940;
      FC_W[31,22] := -0.42096645;
      FC_W[31,23] := -0.97618204;
      FC_W[31,24] := 0.34915537;
      FC_W[31,25] := -1.14380419;
      FC_W[31,26] := -0.40467715;
      FC_W[31,27] := 0.22540230;
      FC_W[31,28] := -0.17240678;
      FC_W[31,29] := -0.31429800;
      FC_W[31,30] := 0.09541429;
      FC_W[31,31] := 0.13256650;
      FC_W[32,0] := 0.72904527;
      FC_W[32,1] := 0.25362849;
      FC_W[32,2] := 0.18425965;
      FC_W[32,3] := 1.12564695;
      FC_W[32,4] := 1.09717035;
      FC_W[32,5] := -0.10607930;
      FC_W[32,6] := -0.54403681;
      FC_W[32,7] := -0.00028945;
      FC_W[32,8] := 0.35294566;
      FC_W[32,9] := -0.17314267;
      FC_W[32,10] := -0.34798992;
      FC_W[32,11] := -0.87766010;
      FC_W[32,12] := -0.42617315;
      FC_W[32,13] := -0.02681804;
      FC_W[32,14] := 0.11679624;
      FC_W[32,15] := -0.28096551;
      FC_W[32,16] := 1.07819867;
      FC_W[32,17] := -0.05331641;
      FC_W[32,18] := -1.38268411;
      FC_W[32,19] := -0.00677918;
      FC_W[32,20] := 0.12342517;
      FC_W[32,21] := -0.18882462;
      FC_W[32,22] := -0.47358170;
      FC_W[32,23] := -1.19179308;
      FC_W[32,24] := -0.13274875;
      FC_W[32,25] := -0.78998423;
      FC_W[32,26] := -0.06041331;
      FC_W[32,27] := -0.37271225;
      FC_W[32,28] := -0.12921399;
      FC_W[32,29] := -0.04796936;
      FC_W[32,30] := 0.12365351;
      FC_W[32,31] := -0.17588998;
      FC_W[33,0] := 0.01445253;
      FC_W[33,1] := 0.31840366;
      FC_W[33,2] := 0.03322378;
      FC_W[33,3] := 1.49474597;
      FC_W[33,4] := 0.91847956;
      FC_W[33,5] := -0.74406970;
      FC_W[33,6] := -0.78569055;
      FC_W[33,7] := -0.22674447;
      FC_W[33,8] := 0.47290990;
      FC_W[33,9] := -0.15914115;
      FC_W[33,10] := -0.23887566;
      FC_W[33,11] := -0.40964791;
      FC_W[33,12] := -0.72407919;
      FC_W[33,13] := 0.32930201;
      FC_W[33,14] := -0.01322137;
      FC_W[33,15] := -0.37601188;
      FC_W[33,16] := 1.17656970;
      FC_W[33,17] := -0.21293037;
      FC_W[33,18] := -1.84557271;
      FC_W[33,19] := -0.40587011;
      FC_W[33,20] := -0.43811360;
      FC_W[33,21] := -0.20921914;
      FC_W[33,22] := -0.87924773;
      FC_W[33,23] := -1.69527853;
      FC_W[33,24] := 0.01967699;
      FC_W[33,25] := 0.12891591;
      FC_W[33,26] := 0.07191025;
      FC_W[33,27] := -0.87316078;
      FC_W[33,28] := -0.11263954;
      FC_W[33,29] := 0.04022661;
      FC_W[33,30] := 0.25044775;
      FC_W[33,31] := -0.00872215;
      FC_W[34,0] := 0.08387819;
      FC_W[34,1] := 0.35092643;
      FC_W[34,2] := -0.02049987;
      FC_W[34,3] := 1.03023493;
      FC_W[34,4] := 0.82523310;
      FC_W[34,5] := -0.45566607;
      FC_W[34,6] := -0.76615703;
      FC_W[34,7] := 0.06065202;
      FC_W[34,8] := 0.64416420;
      FC_W[34,9] := -0.41033185;
      FC_W[34,10] := -0.20673469;
      FC_W[34,11] := -0.60855699;
      FC_W[34,12] := -0.73614651;
      FC_W[34,13] := 0.24825446;
      FC_W[34,14] := 0.08419260;
      FC_W[34,15] := -0.38494027;
      FC_W[34,16] := 0.99920011;
      FC_W[34,17] := -0.68467540;
      FC_W[34,18] := -1.48794913;
      FC_W[34,19] := -0.26779562;
      FC_W[34,20] := -0.25243282;
      FC_W[34,21] := -0.18282467;
      FC_W[34,22] := -0.41076231;
      FC_W[34,23] := -1.47210300;
      FC_W[34,24] := 0.04287826;
      FC_W[34,25] := 0.05358190;
      FC_W[34,26] := 0.09971944;
      FC_W[34,27] := -0.87701261;
      FC_W[34,28] := -0.13157769;
      FC_W[34,29] := 0.02527844;
      FC_W[34,30] := 0.32077599;
      FC_W[34,31] := 0.28405723;
      FC_W[35,0] := 1.02642119;
      FC_W[35,1] := 0.15478377;
      FC_W[35,2] := 0.34819487;
      FC_W[35,3] := 1.05463827;
      FC_W[35,4] := 1.08805430;
      FC_W[35,5] := 0.13107304;
      FC_W[35,6] := -0.46483186;
      FC_W[35,7] := 0.08113482;
      FC_W[35,8] := 0.20881900;
      FC_W[35,9] := -0.12320897;
      FC_W[35,10] := -0.55036026;
      FC_W[35,11] := -1.13076138;
      FC_W[35,12] := -0.23920335;
      FC_W[35,13] := -0.17934363;
      FC_W[35,14] := 0.33692238;
      FC_W[35,15] := -0.24215315;
      FC_W[35,16] := 1.17133689;
      FC_W[35,17] := 0.24548963;
      FC_W[35,18] := -1.27551270;
      FC_W[35,19] := 0.09112822;
      FC_W[35,20] := 0.34386498;
      FC_W[35,21] := -0.19498780;
      FC_W[35,22] := -0.54745656;
      FC_W[35,23] := -0.95400840;
      FC_W[35,24] := -0.28342932;
      FC_W[35,25] := -1.17111981;
      FC_W[35,26] := -0.11992850;
      FC_W[35,27] := -0.10002410;
      FC_W[35,28] := -0.11364288;
      FC_W[35,29] := -0.03451003;
      FC_W[35,30] := -0.05162375;
      FC_W[35,31] := -0.40207881;
      FC_W[36,0] := 0.32796329;
      FC_W[36,1] := 0.27471870;
      FC_W[36,2] := -1.60319293;
      FC_W[36,3] := -0.17304431;
      FC_W[36,4] := 0.69085610;
      FC_W[36,5] := 2.00758481;
      FC_W[36,6] := 0.14931142;
      FC_W[36,7] := -0.71524823;
      FC_W[36,8] := -0.43883818;
      FC_W[36,9] := 0.68334842;
      FC_W[36,10] := -0.10357545;
      FC_W[36,11] := -0.80496567;
      FC_W[36,12] := -0.23269740;
      FC_W[36,13] := 2.37379217;
      FC_W[36,14] := -0.21255036;
      FC_W[36,15] := -0.35580319;
      FC_W[36,16] := -0.20978326;
      FC_W[36,17] := -0.75257885;
      FC_W[36,18] := 0.39406699;
      FC_W[36,19] := 0.35401195;
      FC_W[36,20] := -0.11612377;
      FC_W[36,21] := -0.38309497;
      FC_W[36,22] := -0.26544514;
      FC_W[36,23] := 0.09461114;
      FC_W[36,24] := -0.98066765;
      FC_W[36,25] := -3.36738920;
      FC_W[36,26] := -0.09037717;
      FC_W[36,27] := -0.05651590;
      FC_W[36,28] := -0.08136930;
      FC_W[36,29] := -0.17011009;
      FC_W[36,30] := 0.32433066;
      FC_W[36,31] := -0.52236450;
      FC_W[37,0] := 1.11602509;
      FC_W[37,1] := 0.13230686;
      FC_W[37,2] := 0.37556839;
      FC_W[37,3] := 1.03695834;
      FC_W[37,4] := 1.10666728;
      FC_W[37,5] := 0.21455918;
      FC_W[37,6] := -0.44370866;
      FC_W[37,7] := 0.10324943;
      FC_W[37,8] := 0.17795388;
      FC_W[37,9] := -0.11435414;
      FC_W[37,10] := -0.59511447;
      FC_W[37,11] := -1.19604099;
      FC_W[37,12] := -0.19990741;
      FC_W[37,13] := -0.20347713;
      FC_W[37,14] := 0.36628124;
      FC_W[37,15] := -0.23054719;
      FC_W[37,16] := 1.19065332;
      FC_W[37,17] := 0.32953432;
      FC_W[37,18] := -1.23666811;
      FC_W[37,19] := 0.11926023;
      FC_W[37,20] := 0.40122989;
      FC_W[37,21] := -0.20119728;
      FC_W[37,22] := -0.55009973;
      FC_W[37,23] := -0.88431180;
      FC_W[37,24] := -0.32038155;
      FC_W[37,25] := -1.28385925;
      FC_W[37,26] := -0.12808827;
      FC_W[37,27] := -0.02247072;
      FC_W[37,28] := -0.11043635;
      FC_W[37,29] := -0.04277689;
      FC_W[37,30] := -0.09206246;
      FC_W[37,31] := -0.45274305;
      FC_W[38,0] := 0.08833387;
      FC_W[38,1] := 0.17063738;
      FC_W[38,2] := 0.40627080;
      FC_W[38,3] := -0.02820471;
      FC_W[38,4] := 1.01802444;
      FC_W[38,5] := 0.00276110;
      FC_W[38,6] := 0.35920566;
      FC_W[38,7] := 0.61928076;
      FC_W[38,8] := -1.45084202;
      FC_W[38,9] := -0.42651275;
      FC_W[38,10] := 0.79540843;
      FC_W[38,11] := -0.19398673;
      FC_W[38,12] := 0.25156212;
      FC_W[38,13] := -0.66952437;
      FC_W[38,14] := 0.86726129;
      FC_W[38,15] := 2.49315405;
      FC_W[38,16] := -0.92725694;
      FC_W[38,17] := 0.10850580;
      FC_W[38,18] := -1.27549517;
      FC_W[38,19] := 0.11709256;
      FC_W[38,20] := 0.72766936;
      FC_W[38,21] := 0.85779226;
      FC_W[38,22] := -1.21616077;
      FC_W[38,23] := 1.35759783;
      FC_W[38,24] := -2.16640043;
      FC_W[38,25] := 0.38234365;
      FC_W[38,26] := 0.64837205;
      FC_W[38,27] := -1.83503079;
      FC_W[38,28] := 0.13642681;
      FC_W[38,29] := -0.32257289;
      FC_W[38,30] := 0.36630678;
      FC_W[38,31] := 0.58749110;
      FC_W[39,0] := -1.34213960;
      FC_W[39,1] := -0.39452556;
      FC_W[39,2] := 0.05640002;
      FC_W[39,3] := 2.78641391;
      FC_W[39,4] := -0.53834760;
      FC_W[39,5] := 1.18857467;
      FC_W[39,6] := 1.89260530;
      FC_W[39,7] := 0.14089946;
      FC_W[39,8] := 0.45307723;
      FC_W[39,9] := -0.32008633;
      FC_W[39,10] := 1.56231987;
      FC_W[39,11] := -1.36977983;
      FC_W[39,12] := -0.00040331;
      FC_W[39,13] := -0.25972384;
      FC_W[39,14] := 0.55241877;
      FC_W[39,15] := -0.22095785;
      FC_W[39,16] := -0.25172147;
      FC_W[39,17] := 0.70830828;
      FC_W[39,18] := -0.34716275;
      FC_W[39,19] := -0.04873657;
      FC_W[39,20] := 0.35393974;
      FC_W[39,21] := 0.44481412;
      FC_W[39,22] := 0.93055451;
      FC_W[39,23] := 0.49923140;
      FC_W[39,24] := -0.22098441;
      FC_W[39,25] := -0.13471889;
      FC_W[39,26] := 0.40598431;
      FC_W[39,27] := -0.08490270;
      FC_W[39,28] := 0.20210928;
      FC_W[39,29] := 0.73309517;
      FC_W[39,30] := 0.38844252;
      FC_W[39,31] := 0.51791489;
      FC_B[0] := -0.17348060;
      FC_B[1] := -0.21796906;
      FC_B[2] := 0.11251362;
      FC_B[3] := 0.42275771;
      FC_B[4] := -0.31992450;
      FC_B[5] := 0.49974471;
      FC_B[6] := 0.19967580;
      FC_B[7] := 0.00543070;
      FC_B[8] := 0.32960236;
      FC_B[9] := -0.07780683;
      FC_B[10] := -0.24855255;
      FC_B[11] := -0.18560880;
      FC_B[12] := -0.50896728;
      FC_B[13] := -0.23425932;
      FC_B[14] := 0.47963727;
      FC_B[15] := -0.21440034;
      FC_B[16] := 0.07365502;
      FC_B[17] := -0.34304526;
      FC_B[18] := 0.51340127;
      FC_B[19] := -1.11249006;
      FC_B[20] := -0.08351764;
      FC_B[21] := -0.14279529;
      FC_B[22] := -1.24779224;
      FC_B[23] := -0.57185590;
      FC_B[24] := -0.76752335;
      FC_B[25] := -0.77601463;
      FC_B[26] := -1.05892229;
      FC_B[27] := 0.55543548;
      FC_B[28] := 0.56929213;
      FC_B[29] := 0.66746068;
      FC_B[30] := -1.25867748;
      FC_B[31] := -0.60353893;
      FC_B[32] := -0.68596536;
      FC_B[33] := -0.86961538;
      FC_B[34] := -1.29853678;
      FC_B[35] := -0.29465187;
      FC_B[36] := 0.18345499;
      FC_B[37] := -0.19968984;
      FC_B[38] := 0.11414208;
      FC_B[39] := 1.22691560;

END_DATA_BLOCK
